FUNCTION_BLOCK Status_Remota_HMI (* Service Interface Function Block Type *)
  (* Standard: 61499-2 *)
  (* Version 1.0, 23/10/2026, Hidryco, Hidryco, IHM do Status_Remota *)
  PACKAGE Hidryco.HidrycoLib;
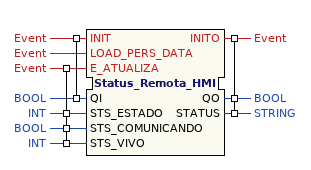
  EVENT_INPUT
    INIT WITH QI;
    LOAD_PERS_DATA; (* Reenvia os parametros persistentes *)
    E_ATUALIZA WITH STS_ESTADO, STS_COMUNICANDO, STS_VIVO; (* Atualizacao de status *)
  END_EVENT
  EVENT_OUTPUT
    INITO WITH QO, STATUS;
  END_EVENT
  VAR_INPUT
    QI : BOOL;
    STS_ESTADO : INT; (* 0 aguardando, 1 comunicando, 2 sem comunicacao *)
    STS_COMUNICANDO : BOOL; (* Remota comunicando *)
    STS_VIVO : INT; (* Sinal de vida (muda a cada 2 s): a IHM acusa CLP sem dados se parar *)
  END_VAR
  VAR_OUTPUT
    QO : BOOL; (* Event Output Qualifier *)
    STATUS : STRING; (* Service Status *)
  END_VAR
  SERVICE /
    SEQUENCE 
    END_SEQUENCE
  END_SERVICE
END_FUNCTION_BLOCK
